Fanuc KAREL source: kt00579.KL

-- PROVISIONAL review KL for V770-1; original PC SHA256 4b285672947085c55b58453ee09e15348cdbb2985152c3257141fc63c5994262
-- Incomplete behavior may be omitted. Consult companion uncertainty JSON. Do not deploy.
PROGRAM KT00579
%NOLOCKGROUP
VAR
  I2 : INTEGER
-- UNRESOLVED_DECL V1 type=000013
-- UNRESOLVED_DECL OUT type=000013
BEGIN
  -- UNRESOLVED_PC offsets 5-20; opcodes 2E,22,32,35
  -- UNRESOLVED_PC offsets 25-36; opcodes 2E,23
  -- UNRESOLVED_PC offsets 41-63; opcodes 49,21,89,4A
  -- UNRESOLVED_PC offsets 68-72; opcodes 7F
END KT00579
